(* IEC 61131-3 sources: trust-platform/examples/OSCAT/battery_energy_storage_facade/oop/src, 3 files *)

(* ---- Main.st ---- *)
(* Record role: BessSnapshot is a deterministic PLC-side record for tests and runtime readers. *)
TYPE BessSnapshot :
STRUCT
    Ready : BOOL;
    StateOfChargePct : REAL;
    PowerCommandKw : REAL;
    AlarmCount : INT;
    FireIsolated : BOOL;
END_STRUCT
END_TYPE

(* Pattern role: IBessAlarmSubscriber is the contract boundary for the Facade and Observer example. *)
INTERFACE IBessAlarmSubscriber
    METHOD OnAlarm
    VAR_INPUT
        AlarmClass : BYTE;
        AlarmCode : WORD;
    END_VAR
    END_METHOD
END_INTERFACE

(* Pattern role: BessHistorianSubscriber is a concrete implementation in the Facade and Observer example. *)
FUNCTION_BLOCK BessHistorianSubscriber IMPLEMENTS IBessAlarmSubscriber
VAR
    AlarmCountValue : INT;
END_VAR
METHOD PUBLIC OnAlarm
VAR_INPUT
    AlarmClass : BYTE;
    AlarmCode : WORD;
END_VAR
AlarmCountValue := AlarmCountValue + INT#1;
END_METHOD
PUBLIC PROPERTY AlarmCount : INT
GET
    AlarmCount := AlarmCountValue;
END_GET
END_PROPERTY
END_FUNCTION_BLOCK

(* Pattern role: BessMqttSubscriber is a concrete implementation in the Facade and Observer example. *)
FUNCTION_BLOCK BessMqttSubscriber IMPLEMENTS IBessAlarmSubscriber
VAR
    PublishReadyValue : BOOL;
END_VAR
METHOD PUBLIC OnAlarm
VAR_INPUT
    AlarmClass : BYTE;
    AlarmCode : WORD;
END_VAR
PublishReadyValue := TRUE;
END_METHOD
PUBLIC PROPERTY PublishReady : BOOL
GET
    PublishReady := PublishReadyValue;
END_GET
END_PROPERTY
END_FUNCTION_BLOCK

(* Composition role: BessAlarmBus owns the collaborating objects used by this Facade and Observer example. *)
FUNCTION_BLOCK BessAlarmBus
VAR
    Historian : IBessAlarmSubscriber;
    Mqtt : IBessAlarmSubscriber;
END_VAR
METHOD PUBLIC Subscribe
VAR_INPUT
    HistorianSub : IBessAlarmSubscriber;
    MqttSub : IBessAlarmSubscriber;
END_VAR
Historian := HistorianSub;
Mqtt := MqttSub;
END_METHOD
METHOD PUBLIC Publish
VAR_INPUT
    AlarmClass : BYTE;
    AlarmCode : WORD;
END_VAR
Historian.OnAlarm(AlarmClass := AlarmClass, AlarmCode := AlarmCode);
Mqtt.OnAlarm(AlarmClass := AlarmClass, AlarmCode := AlarmCode);
END_METHOD
END_FUNCTION_BLOCK

(* Composition role: BatteryRack owns the collaborating objects used by this Facade and Observer example. *)
FUNCTION_BLOCK BatteryRack
VAR
    SocValue : REAL;
    TempFilter : Pt1Filter;
END_VAR
METHOD PUBLIC Initialize
TempFilter.Initialize();
TempFilter.Configure(TimeConstant := T#2s, Gain := REAL#1.0);
END_METHOD
METHOD PUBLIC Update
VAR_INPUT
    StateOfChargePct : REAL;
END_VAR
SocValue := LIMIT(REAL#0.0, StateOfChargePct, REAL#100.0);
END_METHOD
PUBLIC PROPERTY StateOfChargePct : REAL
GET
    StateOfChargePct := SocValue;
END_GET
END_PROPERTY
END_FUNCTION_BLOCK

(* Composition role: InverterUnit owns the collaborating objects used by this Facade and Observer example. *)
FUNCTION_BLOCK InverterUnit
VAR
    EnabledValue : BOOL;
    PowerCommandValue : REAL;
END_VAR
METHOD PUBLIC Command
VAR_INPUT
    Enabled : BOOL;
    PowerKw : REAL;
END_VAR
EnabledValue := Enabled;
IF Enabled THEN
    PowerCommandValue := LIMIT(REAL#-250.0, PowerKw, REAL#250.0);
ELSE
    PowerCommandValue := REAL#0.0;
END_IF;
END_METHOD
PUBLIC PROPERTY PowerCommandKw : REAL
GET
    PowerCommandKw := PowerCommandValue;
END_GET
END_PROPERTY
PUBLIC PROPERTY Enabled : BOOL
GET
    Enabled := EnabledValue;
END_GET
END_PROPERTY
END_FUNCTION_BLOCK

(* Composition role: EnergyStorageCabinet owns the collaborating objects used by this Facade and Observer example. *)
FUNCTION_BLOCK EnergyStorageCabinet
VAR
    Rack : BatteryRack;
    Inverter : InverterUnit;
    AlarmBus : BessAlarmBus;
    Historian : BessHistorianSubscriber;
    Mqtt : BessMqttSubscriber;
    EnabledValue : BOOL;
    SnapshotValue : BessSnapshot;
END_VAR

METHOD PUBLIC Initialize
Rack.Initialize();
AlarmBus.Subscribe(HistorianSub := Historian, MqttSub := Mqtt);
END_METHOD

METHOD PUBLIC Enable
EnabledValue := TRUE;
END_METHOD

METHOD PUBLIC Disable
EnabledValue := FALSE;
Inverter.Command(Enabled := FALSE, PowerKw := REAL#0.0);
END_METHOD

METHOD PUBLIC Update : BessSnapshot
VAR_INPUT
    StateOfChargePct : REAL;
    GridPowerCommandKw : REAL;
    FireInputHealthy : BOOL;
END_VAR
Rack.Update(StateOfChargePct := StateOfChargePct);
SnapshotValue.StateOfChargePct := Rack.StateOfChargePct;
IF NOT FireInputHealthy THEN
    Disable();
    SnapshotValue.FireIsolated := TRUE;
    AlarmBus.Publish(AlarmClass := BYTE#3, AlarmCode := WORD#16#A701);
ELSE
    SnapshotValue.FireIsolated := FALSE;
    Inverter.Command(Enabled := EnabledValue, PowerKw := GridPowerCommandKw);
END_IF;
SnapshotValue.Ready := EnabledValue AND FireInputHealthy;
SnapshotValue.PowerCommandKw := Inverter.PowerCommandKw;
SnapshotValue.AlarmCount := Historian.AlarmCount;
Update := SnapshotValue;
END_METHOD

METHOD PUBLIC Snapshot : BessSnapshot
Snapshot := SnapshotValue;
END_METHOD

PUBLIC PROPERTY StateOfChargePct : REAL
GET
    StateOfChargePct := SnapshotValue.StateOfChargePct;
END_GET
END_PROPERTY
PUBLIC PROPERTY PowerCommandKw : REAL
GET
    PowerCommandKw := SnapshotValue.PowerCommandKw;
END_GET
END_PROPERTY
PUBLIC PROPERTY AlarmCount : INT
GET
    AlarmCount := SnapshotValue.AlarmCount;
END_GET
END_PROPERTY
PUBLIC PROPERTY FireIsolated : BOOL
GET
    FireIsolated := SnapshotValue.FireIsolated;
END_GET
END_PROPERTY
PUBLIC PROPERTY MqttPublishReady : BOOL
GET
    MqttPublishReady := Mqtt.PublishReady;
END_GET
END_PROPERTY
END_FUNCTION_BLOCK

(* Scan role: Main wires the example objects and exposes the PLC call path under test. *)
PROGRAM Main
VAR
    Cabinet : EnergyStorageCabinet;
    EnableCommand : BOOL;
    FireInputHealthy : BOOL;
    SocRaw : INT;
    GridCommandRaw : INT;
    Snapshot : BessSnapshot;
    InverterEnableOut : BOOL;
    FireIsolateOut : BOOL;
END_VAR
Cabinet.Initialize();
IF EnableCommand THEN
    Cabinet.Enable();
END_IF;
Snapshot := Cabinet.Update(StateOfChargePct := INT_TO_REAL(SocRaw), GridPowerCommandKw := INT_TO_REAL(GridCommandRaw), FireInputHealthy := FireInputHealthy);
InverterEnableOut := Snapshot.Ready;
FireIsolateOut := Snapshot.FireIsolated;
END_PROGRAM

(* ---- Configuration.st ---- *)
CONFIGURATION BatteryEnergyStorageFacadeOopConfiguration
RESOURCE Cpu0 ON PLC
    TASK MainTask (INTERVAL := T#100ms, PRIORITY := 1);
    PROGRAM Cabinet WITH MainTask : Main;
END_RESOURCE
VAR_CONFIG
    Cabinet.EnableCommand AT %IX0.0 : BOOL;
    Cabinet.FireInputHealthy AT %IX0.1 : BOOL;
    Cabinet.SocRaw AT %IW0 : INT;
    Cabinet.GridCommandRaw AT %IW2 : INT;
    Cabinet.InverterEnableOut AT %QX0.0 : BOOL;
    Cabinet.FireIsolateOut AT %QX0.1 : BOOL;
END_VAR
END_CONFIGURATION

(* ---- Tests.st ---- *)
TEST_PROGRAM BessFacadeExposesCabinetSnapshot
VAR
    Cabinet : EnergyStorageCabinet;
    Snapshot : BessSnapshot;
END_VAR
Cabinet.Initialize();
Cabinet.Enable();
Snapshot := Cabinet.Update(StateOfChargePct := REAL#70.0, GridPowerCommandKw := REAL#120.0, FireInputHealthy := TRUE);
ASSERT_TRUE(IN := Snapshot.Ready);
ASSERT_NEAR(EXPECTED := REAL#120.0, ACTUAL := Snapshot.PowerCommandKw, DELTA := REAL#0.001);
END_TEST_PROGRAM

TEST_PROGRAM BessObserverPublishesFireAlarm
VAR
    Cabinet : EnergyStorageCabinet;
    Snapshot : BessSnapshot;
END_VAR
Cabinet.Initialize();
Cabinet.Enable();
Snapshot := Cabinet.Update(StateOfChargePct := REAL#70.0, GridPowerCommandKw := REAL#120.0, FireInputHealthy := FALSE);
ASSERT_TRUE(IN := Snapshot.FireIsolated);
ASSERT_EQUAL(EXPECTED := INT#1, ACTUAL := Snapshot.AlarmCount);
ASSERT_TRUE(IN := Cabinet.MqttPublishReady);
END_TEST_PROGRAM

(* Multi-scan facade lifecycle test: drives the cabinet through enable,
   alarm trip, and disable on one instance. Catches bugs where Enable/
   Disable state leaks across scans, where the snapshot freezes after
   the first call, or where Disable doesn't actually zero the power
   command. *)
TEST_PROGRAM BessFacadeLifecycleTracksEnableDisableAcrossScans
VAR
    Cabinet : EnergyStorageCabinet;
    SnapshotEnabled : BessSnapshot;
    SnapshotAlarmed : BessSnapshot;
    SnapshotDisabled : BessSnapshot;
END_VAR

Cabinet.Initialize();
Cabinet.Enable();

(* Scan 1: healthy, command honored *)
SnapshotEnabled := Cabinet.Update(StateOfChargePct := REAL#70.0, GridPowerCommandKw := REAL#100.0, FireInputHealthy := TRUE);
ASSERT_TRUE(IN := SnapshotEnabled.Ready);

(* Scan 2: fire input fails, cabinet must isolate *)
SnapshotAlarmed := Cabinet.Update(StateOfChargePct := REAL#70.0, GridPowerCommandKw := REAL#100.0, FireInputHealthy := FALSE);
ASSERT_TRUE(IN := SnapshotAlarmed.FireIsolated);

(* Scan 3: explicitly disabled - cabinet stops regardless of command *)
Cabinet.Disable();
SnapshotDisabled := Cabinet.Update(StateOfChargePct := REAL#70.0, GridPowerCommandKw := REAL#100.0, FireInputHealthy := TRUE);
ASSERT_FALSE(IN := SnapshotDisabled.Ready);
ASSERT_NEAR(EXPECTED := REAL#0.0, ACTUAL := SnapshotDisabled.PowerCommandKw, DELTA := REAL#0.001);
END_TEST_PROGRAM

(* Inverter power-command boundary regression: the inverter clamps to
   [-250, 250] kW. Test off-by-one at each rail and beyond. *)
TEST_PROGRAM BessInverterClampsPowerCommandAtRails
VAR
    Cabinet : EnergyStorageCabinet;
    Snapshot : BessSnapshot;
END_VAR
Cabinet.Initialize();
Cabinet.Enable();

(* Just below positive rail: pass-through *)
Snapshot := Cabinet.Update(StateOfChargePct := REAL#50.0, GridPowerCommandKw := REAL#249.9, FireInputHealthy := TRUE);
ASSERT_NEAR(EXPECTED := REAL#249.9, ACTUAL := Snapshot.PowerCommandKw, DELTA := REAL#0.001);

(* At positive rail: pass-through *)
Snapshot := Cabinet.Update(StateOfChargePct := REAL#50.0, GridPowerCommandKw := REAL#250.0, FireInputHealthy := TRUE);
ASSERT_NEAR(EXPECTED := REAL#250.0, ACTUAL := Snapshot.PowerCommandKw, DELTA := REAL#0.001);

(* Above positive rail: clamps to 250 *)
Snapshot := Cabinet.Update(StateOfChargePct := REAL#50.0, GridPowerCommandKw := REAL#500.0, FireInputHealthy := TRUE);
ASSERT_NEAR(EXPECTED := REAL#250.0, ACTUAL := Snapshot.PowerCommandKw, DELTA := REAL#0.001);

(* At negative rail: pass-through *)
Snapshot := Cabinet.Update(StateOfChargePct := REAL#50.0, GridPowerCommandKw := REAL#-250.0, FireInputHealthy := TRUE);
ASSERT_NEAR(EXPECTED := REAL#-250.0, ACTUAL := Snapshot.PowerCommandKw, DELTA := REAL#0.001);

(* Below negative rail: clamps to -250 *)
Snapshot := Cabinet.Update(StateOfChargePct := REAL#50.0, GridPowerCommandKw := REAL#-1000.0, FireInputHealthy := TRUE);
ASSERT_NEAR(EXPECTED := REAL#-250.0, ACTUAL := Snapshot.PowerCommandKw, DELTA := REAL#0.001);
END_TEST_PROGRAM

(* SoC clamp regression: BatteryRack.Update LIMITs SoC to [0, 100]. *)
TEST_PROGRAM BessRackClampsStateOfChargeToValidRange
VAR
    Rack : BatteryRack;
END_VAR
Rack.Initialize();

(* Negative input: clamped to 0 *)
Rack.Update(StateOfChargePct := REAL#-25.0);
ASSERT_NEAR(EXPECTED := REAL#0.0, ACTUAL := Rack.StateOfChargePct, DELTA := REAL#0.001);

(* Above-100 input: clamped to 100 *)
Rack.Update(StateOfChargePct := REAL#150.0);
ASSERT_NEAR(EXPECTED := REAL#100.0, ACTUAL := Rack.StateOfChargePct, DELTA := REAL#0.001);

(* Boundary at 100: pass-through *)
Rack.Update(StateOfChargePct := REAL#100.0);
ASSERT_NEAR(EXPECTED := REAL#100.0, ACTUAL := Rack.StateOfChargePct, DELTA := REAL#0.001);

(* Boundary at 0: pass-through *)
Rack.Update(StateOfChargePct := REAL#0.0);
ASSERT_NEAR(EXPECTED := REAL#0.0, ACTUAL := Rack.StateOfChargePct, DELTA := REAL#0.001);
END_TEST_PROGRAM

(* Per-subscriber isolation: drive the alarm bus directly. Both
   subscribers should fire on every Publish; counts and flags
   accumulate independently. *)
TEST_PROGRAM BessAlarmBusFansOutToAllSubscribers
VAR
    Bus : BessAlarmBus;
    Historian : BessHistorianSubscriber;
    Mqtt : BessMqttSubscriber;
END_VAR
Bus.Subscribe(HistorianSub := Historian, MqttSub := Mqtt);

(* No publishes yet *)
ASSERT_EQUAL(EXPECTED := INT#0, ACTUAL := Historian.AlarmCount);
ASSERT_FALSE(IN := Mqtt.PublishReady);

(* One publish: each subscriber sees it *)
Bus.Publish(AlarmClass := BYTE#1, AlarmCode := WORD#16#0001);
ASSERT_EQUAL(EXPECTED := INT#1, ACTUAL := Historian.AlarmCount);
ASSERT_TRUE(IN := Mqtt.PublishReady);

(* Many publishes: historian counts each, mqtt flag latches *)
Bus.Publish(AlarmClass := BYTE#2, AlarmCode := WORD#16#0002);
Bus.Publish(AlarmClass := BYTE#3, AlarmCode := WORD#16#0003);
ASSERT_EQUAL(EXPECTED := INT#3, ACTUAL := Historian.AlarmCount);
END_TEST_PROGRAM

(* Repeated fire trips on one cabinet: AlarmCount must increment per
   trip, FireIsolated must follow the input. *)
TEST_PROGRAM BessFacadeAlarmCountAccumulatesAcrossFireTrips
VAR
    Cabinet : EnergyStorageCabinet;
    Snapshot : BessSnapshot;
END_VAR
Cabinet.Initialize();
Cabinet.Enable();

(* Healthy scan *)
Snapshot := Cabinet.Update(StateOfChargePct := REAL#50.0, GridPowerCommandKw := REAL#0.0, FireInputHealthy := TRUE);
ASSERT_EQUAL(EXPECTED := INT#0, ACTUAL := Snapshot.AlarmCount);

(* First fire trip: count goes to 1 *)
Snapshot := Cabinet.Update(StateOfChargePct := REAL#50.0, GridPowerCommandKw := REAL#0.0, FireInputHealthy := FALSE);
ASSERT_EQUAL(EXPECTED := INT#1, ACTUAL := Snapshot.AlarmCount);

(* Re-enable, healthy, then a second fire trip: count goes to 2 *)
Cabinet.Enable();
Snapshot := Cabinet.Update(StateOfChargePct := REAL#50.0, GridPowerCommandKw := REAL#0.0, FireInputHealthy := TRUE);
Snapshot := Cabinet.Update(StateOfChargePct := REAL#50.0, GridPowerCommandKw := REAL#0.0, FireInputHealthy := FALSE);
ASSERT_EQUAL(EXPECTED := INT#2, ACTUAL := Snapshot.AlarmCount);

(* Third trip without re-enable: still triggers a publish (Disable was already true but fire still latches) *)
Snapshot := Cabinet.Update(StateOfChargePct := REAL#50.0, GridPowerCommandKw := REAL#0.0, FireInputHealthy := FALSE);
ASSERT_EQUAL(EXPECTED := INT#3, ACTUAL := Snapshot.AlarmCount);
ASSERT_TRUE(IN := Snapshot.FireIsolated);
END_TEST_PROGRAM

(* Inverter without enable: any command rounds to zero. *)
TEST_PROGRAM BessInverterRequiresEnableForPowerCommand
VAR
    Inverter : InverterUnit;
END_VAR
(* Disabled: PowerCommandKw is zero regardless of input *)
Inverter.Command(Enabled := FALSE, PowerKw := REAL#100.0);
ASSERT_NEAR(EXPECTED := REAL#0.0, ACTUAL := Inverter.PowerCommandKw, DELTA := REAL#0.001);
ASSERT_FALSE(IN := Inverter.Enabled);

(* Enabled: command honored *)
Inverter.Command(Enabled := TRUE, PowerKw := REAL#100.0);
ASSERT_NEAR(EXPECTED := REAL#100.0, ACTUAL := Inverter.PowerCommandKw, DELTA := REAL#0.001);
ASSERT_TRUE(IN := Inverter.Enabled);

(* Disable again: drops to zero on next call *)
Inverter.Command(Enabled := FALSE, PowerKw := REAL#100.0);
ASSERT_NEAR(EXPECTED := REAL#0.0, ACTUAL := Inverter.PowerCommandKw, DELTA := REAL#0.001);
END_TEST_PROGRAM
